(* IEC 61131-3 sources: plc-iiot-stack/src/DUTs/Iiot, 21 files *)

(* ---- E_IiotAlarmPriority.dut.st ---- *)
// Назначение: приоритет тревоги (коды PL.E_AlarmPriority).
// Документ:   docs/plc_mqtt.md
{attribute 'qualified_only'}
{attribute 'strict'}
TYPE E_IiotAlarmPriority :
(
    None := 0,   // выключена
    Low := 1,   // 'Low'
    Medium := 2,   // 'Medium'
    High := 3,   // 'High'
    Critical := 4   // 'Critical'
) INT;
END_TYPE

(* ---- E_IiotAlarmReason.dut.st ---- *)
// Назначение: причина события тревоги (коды PL.E_AlarmEventReason).
// Документ:   docs/plc_mqtt.md
{attribute 'qualified_only'}
{attribute 'strict'}
TYPE E_IiotAlarmReason :
(
    None := 0,   // нет
    Activated := 1,   // условие появилось
    Cleared := 2,   // условие ушло
    Acked := 3,   // квитирована
    Shelved := 4,   // отложена
    Unshelved := 5,   // возвращена командой
    ShelveExpired := 6,   // возвращена по таймауту
    Suppressed := 7,   // подавлена
    Unsuppressed := 8,   // подавление снято
    OosOn := 9,   // выведена из работы
    OosOff := 10   // введена в работу
) INT;
END_TYPE

(* ---- E_IiotAlarmState.dut.st ---- *)
// Назначение: состояние тревоги (коды PL.E_AlarmState).
// Документ:   docs/plc_mqtt.md
{attribute 'qualified_only'}
{attribute 'strict'}
TYPE E_IiotAlarmState :
(
    Normal := 0,   // норма
    ActiveUnack := 1,   // активна, не квитирована
    ActiveAck := 2,   // активна, квитирована
    RtnUnack := 3,   // вернулась в норму без квитирования
    Shelved := 4,   // отложена
    SuppressedByDesign := 5,   // подавлена логикой
    OutOfService := 6   // выведена из работы с устройством
) INT;
END_TYPE

(* ---- E_IiotCmdKind.dut.st ---- *)
// Назначение: вид команды по полю value (command.schema.json).
// Документ:   docs/plc_mqtt.md
{attribute 'qualified_only'}
{attribute 'strict'}
TYPE E_IiotCmdKind :
(
    Pulse := 0,   // импульс: поля value быть не должно
    Value := 1,   // значение: value обязательно (SpeedSp, SubstValue)
    Mask := 2   // маска: value — целое 0..65535 (AckReq, ShelveReq, UnshelveReq)
) INT;
END_TYPE

(* ---- E_IiotCmdReason.dut.st ---- *)
// Назначение: причина в ответе на команду (поле reason, data_schema 5.1).
// Документ:   docs/plc_mqtt.md
{attribute 'qualified_only'}
{attribute 'strict'}
TYPE E_IiotCmdReason :
(
    Ok := 0,   // 'ok': принята (result = accepted)
    NotWhitelisted := 1,   // 'not_whitelisted': пары (устройство, команда) нет в белом списке
    OutOfRange := 2,   // 'out_of_range': value вне [min; max]
    InvalidPayload := 3,   // 'invalid_payload': не по command.schema.json
    UnsupportedVersion := 4,   // 'unsupported_version': мажорная версия не 1
    TopicMismatch := 5,   // 'topic_mismatch': command в теле не совпадает с топиком
    Retained := 6,   // 'retained': сообщение с флагом retain
    Expired := 7,   // 'expired': ts дальше допуска от часов ПЛК (или часов нет)
    Duplicate := 8,   // 'duplicate': cmd_id среди последних 16
    RateLimited := 9,   // 'rate_limited': больше 10 команд за 10 с
    DeviceRejected := 10,   // 'device_rejected': устройство отказало (cmd_result)
    Timeout := 11   // 'timeout': устройство не обработало команду
) INT;
END_TYPE

(* ---- E_IiotCommand.dut.st ---- *)
// Назначение: команда (поле command и последний уровень топика): имя поля ST_<Dev>Cmd устройства или
//             ST_StationCmd станции флагмана.
// Документ:   docs/plc_mqtt.md
{attribute 'qualified_only'}
{attribute 'strict'}
TYPE E_IiotCommand :
(
    None := 0,   // не распознана
    SetAuto := 1,   // stCommon.xSetAuto
    SetManual := 2,   // stCommon.xSetManual
    SetOos := 3,   // stCommon.xSetOos
    Start := 4,   // xStart
    Stop := 5,   // xStop
    SpeedSp := 6,   // rSpeedSp_pct: значение 0..100 %
    ResetMaint := 7,   // xResetMaint
    SubstValue := 8,   // rSubstValue_eu / xSubstValue: значение
    Ack := 9,   // stCommon.xAck
    Reset := 10,   // stCommon.xReset
    AckReq := 11,   // stCommon.wAckReq: маска 0..65535
    ShelveReq := 12,   // stCommon.wShelveReq: маска
    UnshelveReq := 13,   // stCommon.wUnshelveReq: маска
    SetStepped := 14,   // станция: xSetStepped
    SetLevelPid := 15,   // станция: xSetLevelPid
    AckAll := 16,   // станция: xAckAll
    ResetAll := 17,   // станция: xResetAll
    Silence := 18   // станция: xSilence
) INT;
END_TYPE

(* ---- E_IiotNe107.dut.st ---- *)
// Назначение: сводный статус связи в духе NAMUR NE 107 (те же коды, что PL.E_Ne107Status флагмана).
// Документ:   docs/plc_mqtt.md
{attribute 'qualified_only'}
{attribute 'strict'}
TYPE E_IiotNe107 :
(
    Good := 0,   // норма: связь есть, публикации проходят
    MaintenanceRequired := 1,   // M: связь есть, но публикации отклоняются (очередь клиента)
    OutOfSpecification := 2,   // S: связь потеряна или не установлена, идут повторы
    CheckFunction := 3,   // C: обмен выключен, нет часов или первое подключение
    Failure := 4   // F: подряд неудачных подключений не меньше порога
) INT;
END_TYPE

(* ---- E_IiotQuality.dut.st ---- *)
// Назначение: качество значения телеметрии (поле quality, data_schema 3.2).
// Документ:   docs/plc_mqtt.md
{attribute 'qualified_only'}
{attribute 'strict'}
TYPE E_IiotQuality :
(
    Good := 0,   // 'good': Good или MaintenanceRequired, значение достоверно
    Uncertain := 1,   // 'uncertain': CheckFunction или OutOfSpecification
    Bad := 2   // 'bad': Failure, недостоверное значение, нет связи с ПЧ
) INT;
END_TYPE

(* ---- E_IiotValueKind.dut.st ---- *)
// Назначение: вид значения метрики в JSON.
// Документ:   docs/plc_mqtt.md
{attribute 'qualified_only'}
{attribute 'strict'}
TYPE E_IiotValueKind :
(
    Analog := 0,   // число с дробной частью: analog и накопительные REAL (наработка)
    Integer := 1   // целое: discrete (0/1), enum (код), counter, integer
) INT;
END_TYPE

(* ---- E_MqttConnState.dut.st ---- *)
// Назначение: состояние связи с брокером (FB_MqttDiag).
// Документ:   docs/plc_mqtt.md
{attribute 'qualified_only'}
{attribute 'strict'}
TYPE E_MqttConnState :
(
    Disabled := 0,   // обмен выключен (xEnable = FALSE) или нет часов
    Connecting := 1,   // подключение запрошено, ждём
    Connected := 2,   // связь есть
    Backoff := 3,   // пауза перед повторным подключением
    Closing := 4   // штатное отключение: опубликовано offline/shutdown, следующий вызов — разрыв
) INT;
END_TYPE

(* ---- E_MqttQos.dut.st ---- *)
// Назначение: уровень качества обслуживания MQTT (QoS).
// Документ:   docs/plc_mqtt.md
{attribute 'qualified_only'}
{attribute 'strict'}
TYPE E_MqttQos :
(
    AtMostOnce := 0,   // QoS 0: не более одного раза
    AtLeastOnce := 1,   // QoS 1: не менее одного раза (возможны повторы)
    ExactlyOnce := 2   // QoS 2: ровно один раз
) INT;
END_TYPE

(* ---- ST_IiotAlarm.dut.st ---- *)
// Назначение: тревога: настройка, текущее и последнее опубликованное состояние.
// Документ:   docs/plc_mqtt.md
{attribute 'qualified_only'}
TYPE ST_IiotAlarm :
STRUCT
    stCfg : ST_IiotAlarmCfg;
    eState : E_IiotAlarmState := E_IiotAlarmState.Normal;       // по словам устройства
    eLastState : E_IiotAlarmState := E_IiotAlarmState.Normal;   // последнее опубликованное
    xSent : BOOL;                                                // опубликовано с последнего подключения
    // Последняя публикация (ts и prev_state): после переподключения она повторяется без изменений —
    // в InfluxDB это та же точка, а не новое срабатывание. 0 — с запуска ПЛК не публиковалась.
    uliEventTs_ms : ULINT;
    eEventPrev : E_IiotAlarmState := E_IiotAlarmState.Normal;
END_STRUCT
END_TYPE

(* ---- ST_IiotAlarmCfg.dut.st ---- *)
// Назначение: тревога перечня флагмана (scada_alarms.csv, station_alarms.csv): номер, источник, суффикс,
//             бит в словах тревог, приоритет.
// Документ:   docs/plc_mqtt.md
{attribute 'qualified_only'}
TYPE ST_IiotAlarmCfg :
STRUCT
    udiId : UDINT;                                   // устройство: dev_no * 10 + слот; станция: 100000 + slot
    sDevice : STRING(GVL_Const.IIOT_DEVICE_LEN);     // 'P101', 'KNS1'
    sSuffix : STRING(GVL_Const.IIOT_SUFFIX_LEN);     // 'FTS'; код тревоги — <sDevice>.<sSuffix>
    uiSlot : UINT;                                   // бит в словах тревог (у станции slot - 1)
    ePriority : E_IiotAlarmPriority := E_IiotAlarmPriority.Medium;
    diWords : DINT;                                  // строка таблицы слов устройства (ST_IiotAlarmWords)
END_STRUCT
END_TYPE

(* ---- ST_IiotAlarmWords.dut.st ---- *)
// Назначение: слова тревог источника (stSts.stCommon устройства или stStationSts станции) и признак
//             вывода из работы.
// Документ:   docs/plc_mqtt.md
{attribute 'qualified_only'}
TYPE ST_IiotAlarmWords :
STRUCT
    wActive : WORD;          // wAlmActive
    wUnack : WORD;           // wAlmUnack
    wShelved : WORD;         // wAlmShelved: отложен оператором (у станции — и подавлен, и выведен)
    wSuppressed : WORD;      // wAlmSuppressed: подавлен логикой (SuppressedByDesign); у станции 0
    xOutOfService : BOOL;    // eMode = OutOfService
END_STRUCT
END_TYPE

(* ---- ST_IiotCfg.dut.st ---- *)
// Назначение: настройки ПЛК-части IIoT-стека (GVL_Iiot.stIiotCfg); топики — schema/topics.json.
// Документ:   docs/plc_mqtt.md
{attribute 'qualified_only'}
TYPE ST_IiotCfg :
STRUCT
    xEnable : BOOL;                                    // обмен MQTT включён (по умолчанию выключен до наладки)
    xCommandsEnable : BOOL;                            // приём команд MQTT (по умолчанию выключен)
    sSite : STRING(GVL_Const.IIOT_LEVEL_LEN) := 'vodokanal';
    sArea : STRING(GVL_Const.IIOT_LEVEL_LEN) := 'kns1';
    sUnit : STRING(GVL_Const.IIOT_LEVEL_LEN) := 'station';
    sNode : STRING(GVL_Const.IIOT_DEVICE_LEN) := 'PLC1';  // узел ПЛК: status/connection и метрики PLC1
    sSwVersion : STRING(GVL_Const.IIOT_TEXT_LEN) := '0.1.0';
    tTelemetryPeriod : TIME := GVL_Const.TELEMETRY_PERIOD_DEFAULT;
    stBroker : ST_MqttBrokerCfg;
END_STRUCT
END_TYPE

(* ---- ST_IiotCmd.dut.st ---- *)
// Назначение: команда, прошедшая проверки шлюза (FB_MqttCommands.stCmd).
// Документ:   docs/plc_mqtt.md
{attribute 'qualified_only'}
TYPE ST_IiotCmd :
STRUCT
    diRule : DINT;                                  // строка белого списка
    sDevice : STRING(GVL_Const.IIOT_DEVICE_LEN);
    sCommand : STRING(GVL_Const.IIOT_LEVEL_LEN);    // последний уровень топика
    eCommand : E_IiotCommand := E_IiotCommand.None;
    rValue : REAL;                                  // для команд-значений и масок
    sCmdId : STRING(GVL_Const.CMD_ID_LEN);
END_STRUCT
END_TYPE

(* ---- ST_IiotCmdRule.dut.st ---- *)
// Назначение: строка белого списка команд (command_whitelist.csv).
// Документ:   docs/plc_mqtt.md
{attribute 'qualified_only'}
TYPE ST_IiotCmdRule :
STRUCT
    sDevice : STRING(GVL_Const.IIOT_DEVICE_LEN);    // 'P101'
    eCommand : E_IiotCommand := E_IiotCommand.None;
    xRange : BOOL;                                  // у команды есть диапазон value
    rMin : REAL;
    rMax : REAL;
    diDev : DINT;                                   // номер устройства для FB_IiotKnsMap.DeviceCmdState
END_STRUCT
END_TYPE

(* ---- ST_IiotPoint.dut.st ---- *)
// Назначение: метрика телеметрии: настройка, текущее и последнее опубликованное значение.
// Документ:   docs/plc_mqtt.md
{attribute 'qualified_only'}
TYPE ST_IiotPoint :
STRUCT
    stCfg : ST_IiotPointCfg;
    // текущее (заполняет FB_IiotKnsMap.FillPoints или PRG_Iiot)
    lrValue : LREAL;
    eQuality : E_IiotQuality := E_IiotQuality.Bad;
    // последнее опубликованное (FB_MqttTelemetry)
    lrLastValue : LREAL;
    lrLastFinite : LREAL;                           // последнее опубликованное конечное значение
    eLastQuality : E_IiotQuality := E_IiotQuality.Bad;
    ltLastSent : LTIME;
    xSent : BOOL;                                   // опубликовано с последнего подключения
    xForce : BOOL;                                  // опубликовать независимо от изменения (период)
END_STRUCT
END_TYPE

(* ---- ST_IiotPointCfg.dut.st ---- *)
// Назначение: метрика каталога: топик <prefix>/<sPath>, вид, единица, зона нечувствительности.
// Документ:   docs/plc_mqtt.md
{attribute 'qualified_only'}
TYPE ST_IiotPointCfg :
STRUCT
    sPath : STRING(GVL_Const.IIOT_PATH_LEN);        // device/metric, например 'LT101/level'
    sUnit : STRING(GVL_Const.IIOT_UNIT_LEN);        // единица (ASCII); пусто — поля unit нет
    eKind : E_IiotValueKind := E_IiotValueKind.Integer;
    rDeadband : REAL;                               // зона нечувствительности, ед.; 0 — любое изменение
    uiDecimals : UINT := GVL_Const.JSON_REAL_DECIMALS_DEFAULT;   // знаков после точки (Analog)
    xPeriodicOnly : BOOL;                           // только с контрольной публикацией (uptime)
END_STRUCT
END_TYPE

(* ---- ST_IiotSts.dut.st ---- *)
// Назначение: состояние ПЛК-части IIoT-стека для HMI и SCADA (GVL_Iiot.stIiotSts).
// Документ:   docs/plc_mqtt.md
{attribute 'qualified_only'}
TYPE ST_IiotSts :
STRUCT
    eConnState : E_MqttConnState := E_MqttConnState.Disabled;
    eNe107 : E_IiotNe107 := E_IiotNe107.CheckFunction;
    udiConnects : UDINT;
    udiDisconnects : UDINT;
    udiConnectFailures : UDINT;
    diLastError : DINT;
    udiPublished : UDINT;                     // телеметрия и тревоги, принятые клиентом
    udiPublishFailed : UDINT;                 // клиент не принял (повторится)
    uiQueue : UINT;                           // записей ждут публикации
    udiDropped : UDINT;                       // сообщений отброшено (не поместились, ответ не принят)
    udiCmdAccepted : UDINT;
    udiCmdRejected : UDINT;                   // отказы с ответом и без ответа
    eLastCmdReason : E_IiotCmdReason := E_IiotCmdReason.Ok;
    xClockValid : BOOL;                       // часы ПЛК в диапазоне схемы: обмен разрешён
END_STRUCT
END_TYPE

(* ---- ST_MqttBrokerCfg.dut.st ---- *)
// Назначение: параметры подключения к брокеру MQTT (I_MqttClient.Connect).
// Документ:   docs/plc_mqtt.md
{attribute 'qualified_only'}
TYPE ST_MqttBrokerCfg :
STRUCT
    sHost : STRING(GVL_Const.BROKER_HOST_LEN);            // имя или адрес брокера
    uiPort : UINT := GVL_Const.MQTT_PORT_DEFAULT;         // 1883; с TLS обычно 8883
    xTls : BOOL;                                           // TLS; проверка сертификата — забота адаптера
    sClientId : STRING(GVL_Const.BROKER_CLIENT_ID_LEN) := 'kns1-plc1';
    sUser : STRING(GVL_Const.BROKER_SECRET_LEN);
    {attribute 'symbol' := 'none'}
    sPassword : STRING(GVL_Const.BROKER_SECRET_LEN);      // задаётся при наладке; в git и в OPC UA не попадает
    tKeepAlive : TIME := GVL_Const.KEEPALIVE_DEFAULT;
    xCleanSession : BOOL := TRUE;
    sWillTopic : STRING(GVL_Const.MQTT_TOPIC_LEN);        // LWT: заполняет FB_MqttDiag перед Connect
    sWillPayload : STRING(GVL_Const.BROKER_WILL_LEN);     // LWT: заполняет FB_MqttDiag
    xWillRetain : BOOL := TRUE;
END_STRUCT
END_TYPE
